TYPE ST_BatCmd :		// BMS에 보낼 명령
STRUCT
	eCmd		: E_BatCmd;
	nSeq		: UDINT;		// 명령 번호. 바뀌면 새 명령 → 디스패처가 1회 전송
END_STRUCT
END_TYPE

(* stored: Version 1.1.0.1, ProductVersion 3.1.4024.15
   DUT ST_BatCmd: Id {8c209493-1420-48a3-b486-b9ffd7f4f5b5} *)
